Fanuc KAREL source: kb00079.KL

-- PROVISIONAL review KL for V940-1; original PC SHA256 53ddbd067d106dec3582ee036b37a90ae9c84a75a2055f8add2539b9b181da9d
-- Incomplete behavior may be omitted. Consult companion uncertainty JSON. Do not deploy.
PROGRAM KB00079
%NOLOCKGROUP
BEGIN
  -- V9_ZERO_TABLE_METADATA_HINT layout=0002_ascii; no indexed target words; source/name/runtime held
  -- UNRESOLVED_PC offsets 5-12; opcodes 9D,23
  -- UNRESOLVED_PC offsets 17-24; opcodes 9D,23
  -- UNRESOLVED_PC offsets 29-36; opcodes 9D,23
  -- UNRESOLVED_PC offsets 41-77; opcodes 27,22,22,22,27,9D,31,7E,4A
  -- UNRESOLVED_PC offsets 82-86; opcodes 7F
END KB00079
